Staubli VAL3: utBorder.dtx

public string sBorderColour
public string sBorderSytle
public string sBorderWidth
